// TwinCAT 3 PLC project PLC
// ProgramVersion: 3.1.4026.28
// libraries:
//   Tc2_MC2, * (Beckhoff Automation GmbH)
//   Tc2_Standard, * (Beckhoff Automation GmbH)
//   Tc2_System, * (Beckhoff Automation GmbH)
// project tree:
//   Adapters/Nc/ Axes.TcGVL, DriveAxis_Nc.TcPOU
//   Adapters/Simulation/ Accelerometer_Simulated.TcPOU, DigitalOut_SimulatedLidarPower.TcPOU, Gyro_Simulated.TcPOU, Lidar_Simulated.TcPOU, SimulatorLink.TcPOU
//   App/ MAIN.TcPOU, RobotComposition.TcPOU
//   Contracts/ HmiCommand.TcDUT, HmiCommandCode.TcDUT, HmiStatus.TcDUT, MapInfo.TcDUT, MissionState.TcDUT, RobotHmi.TcGVL, SimulatorCommand.TcDUT, SimulatorFeedback.TcDUT, SimulatorIo.TcGVL
//   Core/ BodyMotion.TcDUT, Constants.TcGVL, HardwareError.TcDUT, LaserScan.TcDUT, Parameters.TcGVL, PlatformKind.TcDUT, Pose2D.TcDUT, Twist.TcDUT, Vector3.TcDUT, WheelSpeeds.TcDUT
//   Hal/ I_Accelerometer.TcIO, I_DigitalOut.TcIO, I_DriveAxis.TcIO, I_Gyro.TcIO, I_Lidar.TcIO, Lidar_Watchdog.TcPOU
//   Localization/ I_PoseSource.TcIO, GyroOdometry.TcPOU, WheelOdometry.TcPOU
//   Mapping/ GridCell.TcDUT, OccupancyGrid.TcPOU
//   Mission/ SweepMission.TcPOU
//   Platform/ DiffDrive.TcPOU, DiffDriveKinematics.TcPOU, I_DifferentialDrive.TcIO
//   / PlcTask.TcTTO
// real-time tasks:
//   TASK PlcTask: cycle T#10ms, priority 20, ADS port 350
// motion (NC):
//   TASK NC-Task 1 SAF: cycle T#2ms, priority 4, ADS port 501
//   TASK NC-Task 1 SVB: cycle T#10ms, priority 8, ADS port 511
//   AXIS LeftWheel (id 1)
//     General: UnitName=m
//     Dynamic: AccelerationMaximum=2, DecelerationMaximum=2, Acceleration=1, Deceleration=1, Jerk=10
//     Velo: Maximum=0.6
//     OtherSettings: AllowMotionCmdToSlave=true
//     encoder EncType=1
//     drive DrvType=5
//       Analog: VeloReferenz=0.6, TorqueSetpointScale=10, ScaleFactorActTorque=0.1
//       TimeComp: TaskDelayCycles=1
//     controller CtrType=1
//       CtrPara: PriorControlFactor=1
//         Observer: BandWidth=20
//   AXIS RightWheel (id 2)
//     General: UnitName=m
//     Dynamic: AccelerationMaximum=2, DecelerationMaximum=2, Acceleration=1, Deceleration=1, Jerk=10
//     Velo: Maximum=0.6
//     OtherSettings: AllowMotionCmdToSlave=true
//     encoder EncType=1
//     drive DrvType=5
//       Analog: VeloReferenz=0.6, TorqueSetpointScale=10, ScaleFactorActTorque=0.1
//       TimeComp: TaskDelayCycles=1
//     controller CtrType=1
//       CtrPara: PriorControlFactor=1
//         Observer: BandWidth=20
// variable links:
//   PLC/PLC Instance <-> NC-Task 1 SAF/Axes/LeftWheel
//     PlcTask Inputs/Axes.leftWheel.NcToPlc <-> Outputs/ToPlc
//     PlcTask Outputs/Axes.leftWheel.PlcToNc <-> Inputs/FromPlc
//   PLC/PLC Instance <-> NC-Task 1 SAF/Axes/RightWheel
//     PlcTask Inputs/Axes.rightWheel.NcToPlc <-> Outputs/ToPlc
//     PlcTask Outputs/Axes.rightWheel.PlcToNc <-> Inputs/FromPlc

CONFIGURATION PLC
    RESOURCE PLC ON TwinCAT3
        TASK PlcTask(INTERVAL := T#10ms, PRIORITY := 20);
        PROGRAM MAIN WITH PlcTask : MAIN;
    END_RESOURCE
END_CONFIGURATION

// ---- Contracts/HmiCommand.TcDUT
TYPE HmiCommand :
STRUCT
	sequence : UDINT;
	code : HmiCommandCode;
	manualTwist : Twist;
	pose : Pose2D;
END_STRUCT
END_TYPE

// ---- Contracts/HmiCommandCode.TcDUT
{attribute 'qualified_only'}
{attribute 'strict'}
TYPE HmiCommandCode :
(
	NONE := 0,
	MANUAL_DRIVE,
	START_MAPPING,
	START_SWEEPING,
	PAUSE,
	RESUME,
	STOP,
	GO_TO_DOCK,
	EMERGENCY_STOP,
	RESET,
	SET_POSE
) INT;
END_TYPE

// ---- Contracts/HmiStatus.TcDUT
TYPE HmiStatus :
STRUCT
	acknowledgedSequence : UDINT;
	missionState : MissionState;
	lastRejection : STRING(80);
	estimatedPose : Pose2D;
	isSimulatorConnected : BOOL;
	isLidarOk : BOOL;
	hasMap : BOOL;
END_STRUCT
END_TYPE

// ---- Contracts/MapInfo.TcDUT
// Det GUI-en trenger for å tegne RobotHmi.mapCells.
TYPE MapInfo :
STRUCT
	// Øker hver gang kartet er endret, så serveren bare henter cellene på nytt når det trengs.
	revision : UDINT;
	cellSizeInM : LREAL;
	// Hjørnet til celle [0, 0] i verden.
	originXInM : LREAL;
	originYInM : LREAL;
	widthInCells : UINT;
	heightInCells : UINT;
	// Hvor mye log-odds én enhet i en celle er. 0.1 betyr at 35 i cella er log-odds 3.5.
	logOddsPerUnit : LREAL;
END_STRUCT
END_TYPE

// ---- Contracts/MissionState.TcDUT
{attribute 'qualified_only'}
{attribute 'strict'}
TYPE MissionState :
(
	IDLE := 0,
	MANUAL,
	MAPPING,
	SWEEPING,
	PAUSED,
	RETURNING_TO_DOCK,
	DOCKED,
	EMERGENCY_STOPPED
) INT;
END_TYPE

// ---- Contracts/SimulatorCommand.TcDUT
TYPE SimulatorCommand :
STRUCT
	version : UDINT;
	cycle : UDINT;
	plcTimeInNs : ULINT;
	// The wheels' actual speed and position, from the NC axes. The simulated wheels run at
	// the speed and are nudged towards the position, so they never drift away from NC.
	leftWheelVelocityInMPerS : LREAL;
	rightWheelVelocityInMPerS : LREAL;
	leftWheelPositionInM : LREAL;
	rightWheelPositionInM : LREAL;
	isLeftDriveEnabled : BOOL;
	isRightDriveEnabled : BOOL;
	isLidarPowered : BOOL;
	estimatedPose : Pose2D;
END_STRUCT
END_TYPE

// ---- Contracts/SimulatorFeedback.TcDUT
TYPE SimulatorFeedback :
STRUCT
	version : UDINT;
	sequence : UDINT;
	timeInNs : ULINT;
	leftWheelAngleInRad : LREAL;
	rightWheelAngleInRad : LREAL;
	leftWheelVelocityInRadPerS : LREAL;
	rightWheelVelocityInRadPerS : LREAL;
	angularRateInRadPerS : Vector3;
	accelerationInMPerS2 : Vector3;
	truePose : Pose2D;
	collided : BOOL;
END_STRUCT
END_TYPE

// ---- Core/BodyMotion.TcDUT
TYPE BodyMotion :
STRUCT
	distanceInM : LREAL;
	headingChangeInRad : LREAL;
END_STRUCT
END_TYPE

// ---- Core/HardwareError.TcDUT
TYPE HardwareError :
STRUCT
	isActive : BOOL;
	id : UDINT;
	text : STRING(80);
END_STRUCT
END_TYPE

// ---- Core/LaserScan.TcDUT
TYPE LaserScan :
STRUCT
	sequence : UDINT;
	startTimestampInNs : ULINT;
	scanDurationInS : REAL;
	angleMinInRad : REAL;
	angleIncrementInRad : REAL;
	count : UINT;
	rangesInM : ARRAY[0..Constants.MAX_SCAN_POINTS - 1] OF REAL;
END_STRUCT
END_TYPE

// ---- Core/PlatformKind.TcDUT
{attribute 'qualified_only'}
{attribute 'strict'}
TYPE PlatformKind :
(
	SIMULATION := 0,
	HARDWARE
);
END_TYPE

// ---- Core/Pose2D.TcDUT
TYPE Pose2D :
STRUCT
	x : LREAL;
	y : LREAL;
	thetaInRad : LREAL;
END_STRUCT
END_TYPE

// ---- Core/Twist.TcDUT
TYPE Twist :
STRUCT
	forwardSpeedInMPerS : LREAL;
	yawRateInRadPerS : LREAL;
END_STRUCT
END_TYPE

// ---- Core/Vector3.TcDUT
TYPE Vector3 :
STRUCT
	x : LREAL;
	y : LREAL;
	z : LREAL;
END_STRUCT
END_TYPE

// ---- Core/WheelSpeeds.TcDUT
TYPE WheelSpeeds :
STRUCT
	leftInMPerS : LREAL;
	rightInMPerS : LREAL;
END_STRUCT
END_TYPE

// ---- Mapping/GridCell.TcDUT
// Én rute i kartet. x teller østover og y nordover fra kartets origo, som i verden.
TYPE GridCell :
STRUCT
	x : DINT;
	y : DINT;
END_STRUCT
END_TYPE

// ---- Adapters/Nc/Axes.TcGVL
{attribute 'qualified_only'}
VAR_GLOBAL
	// Link each one to its NC axis in XAE: the axis, Settings, Link To PLC.
	leftWheel : AXIS_REF;
	rightWheel : AXIS_REF;
END_VAR

// ---- Contracts/RobotHmi.TcGVL
{attribute 'qualified_only'}
VAR_GLOBAL
	command : HmiCommand;
	status : HmiStatus;
	// Kartet PLC-en bygger, for GUI-en. Indeksen er [x, y]; y endrer seg raskest i minnet.
	mapInfo : MapInfo;
	mapCells : ARRAY[0..Constants.MAP_WIDTH_IN_CELLS - 1, 0..Constants.MAP_HEIGHT_IN_CELLS - 1] OF SINT;
END_VAR

// ---- Contracts/SimulatorIo.TcGVL
{attribute 'qualified_only'}
VAR_GLOBAL
	command : SimulatorCommand;
	feedback : SimulatorFeedback;
	scan : LaserScan;
END_VAR

// ---- Core/Constants.TcGVL
{attribute 'qualified_only'}
VAR_GLOBAL CONSTANT
	MAX_SCAN_POINTS : UINT := 1024;
	// Kartet er 256 x 256 ruter. Med 5 cm ruter blir det 12,8 x 12,8 m.
	MAP_WIDTH_IN_CELLS : UINT := 256;
	MAP_HEIGHT_IN_CELLS : UINT := 256;
	// Én enhet i en kartcelle er så mye log-odds.
	MAP_LOG_ODDS_PER_UNIT : LREAL := 0.1;
	SIMULATOR_PROTOCOL_VERSION : UDINT := 4;
	SIMULATOR_TIMEOUT_IN_CYCLES : UDINT := 20;
	LIDAR_TIMEOUT_IN_MS : TIME := T#400MS;
	SIMULATOR_NOT_CONNECTED_ERROR_ID : UDINT := 1001;
	LIDAR_TIMEOUT_ERROR_ID : UDINT := 2001;
	AXIS_NOT_LINKED_ERROR_ID : UDINT := 3001;
END_VAR

// ---- Core/Parameters.TcGVL
{attribute 'qualified_only'}
VAR_GLOBAL PERSISTENT
	platform : PlatformKind := PlatformKind.SIMULATION;
	// Hjulradien ligger i NC-skaleringen av aksene, som går i meter langs hjulbanen.
	trackWidthInM : LREAL := 0.40;
	maxWheelSpeedInMPerS : LREAL := 0.6;
	// Hvor fort hjulene får endre fart. Uten disse bruker NC sine standardverdier, og hjulene
	// stopper fra full fart på et par hundredeler, mye brattere enn en ekte robot tåler uten å skli.
	wheelAccelerationInMPerS2 : LREAL := 1.0;
	wheelJerkInMPerS3 : LREAL := 10.0;
	useGyroForHeading : BOOL := FALSE;
	gyroScale : LREAL := 1.0;

	// Hvor lidaren sitter på roboten, sett fra midt mellom hjulene (x fram, y mot venstre),
	// og hvor mye den er dreid. I simulatoren står den midt mellom hjulene og peker rett fram.
	lidarMountXInM : LREAL := 0.0;
	lidarMountYInM : LREAL := 0.0;
	lidarMountThetaInRad : LREAL := 0.0;

	// Kartet. Origo er hjørnet til celle [0, 0]; med -3.4 dekker kartet en garasje på 6 x 6 m med god margin.
	mapCellSizeInM : LREAL := 0.05;
	mapOriginXInM : LREAL := -3.4;
	mapOriginYInM : LREAL := -3.4;
	// Log-odds i tideler (Constants.MAP_LOG_ODDS_PER_UNIT): treff +0.9, fri -0.4, aldri mer enn ±3.5.
	mapHitLogOdds : SINT := 9;
	mapFreeLogOdds : SINT := -4;
	mapMaxLogOdds : SINT := 35;
END_VAR

// ---- Hal/I_Accelerometer.TcIO
INTERFACE I_Accelerometer

PROPERTY AccelerationInMPerS2 : Vector3
GET
END_GET
END_PROPERTY

PROPERTY TimestampInNs : ULINT
GET
END_GET
END_PROPERTY

PROPERTY IsValid : BOOL
GET
END_GET
END_PROPERTY

END_INTERFACE

// ---- Hal/I_DigitalOut.TcIO
INTERFACE I_DigitalOut

METHOD SwitchOn
END_METHOD

METHOD SwitchOff
END_METHOD

PROPERTY IsOn : BOOL
GET
END_GET
END_PROPERTY

END_INTERFACE

// ---- Hal/I_DriveAxis.TcIO
INTERFACE I_DriveAxis

METHOD Execute
END_METHOD

METHOD Enable
END_METHOD

METHOD Disable
END_METHOD

METHOD SetVelocity
VAR_INPUT
	velocityInMPerS : LREAL;
END_VAR
END_METHOD

METHOD TryReset : BOOL
END_METHOD

PROPERTY PositionInM : LREAL
GET
END_GET
END_PROPERTY

PROPERTY VelocityInMPerS : LREAL
GET
END_GET
END_PROPERTY

PROPERTY IsReady : BOOL
GET
END_GET
END_PROPERTY

PROPERTY IsStandingStill : BOOL
GET
END_GET
END_PROPERTY

PROPERTY Error : HardwareError
GET
END_GET
END_PROPERTY

END_INTERFACE

// ---- Hal/I_Gyro.TcIO
INTERFACE I_Gyro

METHOD StartBiasCalibration
END_METHOD

PROPERTY YawRateInRadPerS : LREAL
GET
END_GET
END_PROPERTY

PROPERTY AngularRateInRadPerS : Vector3
GET
END_GET
END_PROPERTY

PROPERTY TimestampInNs : ULINT
GET
END_GET
END_PROPERTY

PROPERTY IsValid : BOOL
GET
END_GET
END_PROPERTY

END_INTERFACE

// ---- Hal/I_Lidar.TcIO
INTERFACE I_Lidar

METHOD Start
END_METHOD

METHOD Stop
END_METHOD

METHOD TryGetScan : BOOL
VAR_INPUT
	scan : REFERENCE TO LaserScan;
END_VAR
END_METHOD

PROPERTY IsRunning : BOOL
GET
END_GET
END_PROPERTY

PROPERTY Error : HardwareError
GET
END_GET
END_PROPERTY

END_INTERFACE

// ---- Localization/I_PoseSource.TcIO
INTERFACE I_PoseSource

METHOD Reset
VAR_INPUT
	pose : Pose2D;
END_VAR
END_METHOD

PROPERTY Pose : Pose2D
GET
END_GET
END_PROPERTY

END_INTERFACE

// ---- Platform/I_DifferentialDrive.TcIO
INTERFACE I_DifferentialDrive

METHOD Execute
END_METHOD

METHOD Enable
END_METHOD

METHOD Disable
END_METHOD

METHOD SetTwist
VAR_INPUT
	desiredTwist : Twist;
END_VAR
END_METHOD

PROPERTY LeftWheelPositionInM : LREAL
GET
END_GET
END_PROPERTY

PROPERTY RightWheelPositionInM : LREAL
GET
END_GET
END_PROPERTY

PROPERTY IsReady : BOOL
GET
END_GET
END_PROPERTY

PROPERTY IsStandingStill : BOOL
GET
END_GET
END_PROPERTY

END_INTERFACE

// ---- App/MAIN.TcPOU
PROGRAM MAIN
VAR
	robot : RobotComposition;
END_VAR

robot.Execute();

END_PROGRAM

// ---- App/RobotComposition.TcPOU
{attribute 'linkalways'}
{attribute 'no_explicit_call' := 'Use the methods of this class'}
{attribute 'enable_dynamic_creation'}
FUNCTION_BLOCK RobotComposition
VAR
	simulator : SimulatorLink;
	leftAxis : DriveAxis_Nc(ncAxis := Axes.leftWheel);
	rightAxis : DriveAxis_Nc(ncAxis := Axes.rightWheel);
	simulatedGyro : Gyro_Simulated(simulator := simulator);
	simulatedAccelerometer : Accelerometer_Simulated(simulator := simulator);
	simulatedLidar : Lidar_Simulated(simulator := simulator);
	simulatedLidarPower : DigitalOut_SimulatedLidarPower;

	gyro : I_Gyro;
	accelerometer : I_Accelerometer;
	lidarPower : I_DigitalOut;
	lidar : Lidar_Watchdog;
	drive : DiffDrive;
	odometry : WheelOdometry;
	gyroOdometry : GyroOdometry;
	grid : OccupancyGrid;
	mission : SweepMission;

	scan : LaserScan;
	requestedPose : Pose2D;
	isInitialized : BOOL;
END_VAR

METHOD Execute
IF NOT isInitialized THEN
	Initialize();
END_IF

IF Parameters.platform = PlatformKind.SIMULATION THEN
	simulator.Execute();
END_IF

lidar.Execute();
IF lidar.TryGetScan(scan) AND mission.State = MissionState.MAPPING THEN
	// Kommer i M4: scan matching, som retter posisjonen mot kartet før scannet legges inn.
	grid.Integrate(scan := scan, pose := EstimatedPose());
	grid.Publish(RobotHmi.mapInfo, RobotHmi.mapCells);
END_IF

odometry.Execute();
gyroOdometry.Execute();
mission.Execute();
IF mission.TryTakePoseRequest(requestedPose) THEN
	odometry.Reset(requestedPose);
	gyroOdometry.Reset(requestedPose);
END_IF
IF mission.TryTakeMapClearRequest() THEN
	grid.Clear();
	grid.Publish(RobotHmi.mapInfo, RobotHmi.mapCells);
END_IF

IF mission.ShouldDrive THEN
	drive.Enable();
	drive.SetTwist(mission.DesiredTwist);
ELSE
	drive.Disable();
END_IF
drive.Execute();

IF Parameters.platform = PlatformKind.SIMULATION THEN
	SendWheelsToSimulator();
END_IF

PublishStatus();
END_METHOD

METHOD PRIVATE Initialize
VAR
	start : Pose2D;
END_VAR
CASE Parameters.platform OF
	PlatformKind.SIMULATION:
		gyro := simulatedGyro;
		accelerometer := simulatedAccelerometer;
		lidar.Wrap(simulatedLidar);
		lidarPower := simulatedLidarPower;
	PlatformKind.HARDWARE:
		// Kommer i M7: Gyro_EP3751 og valgt LIDAR-adapter. Hjulene bruker de samme NC-aksene.
		RETURN;
END_CASE

drive.Connect(leftAxis, rightAxis);

lidarPower.SwitchOn();
lidar.Start();
odometry.Connect(drive);
odometry.Reset(start);
gyroOdometry.Connect(drive, gyro);
gyroOdometry.Reset(start);
grid.Clear();
grid.Publish(RobotHmi.mapInfo, RobotHmi.mapCells);
isInitialized := TRUE;
END_METHOD

METHOD PRIVATE SendWheelsToSimulator
// I simuleringen er NC-aksene motor og enkoder. Simulatoren får vite hvor langt hjulene faktisk har gått,
// lar de simulerte hjulene følge det nøyaktig, og flytter roboten etter det, med sluring og kollisjoner.
SimulatorIo.command.leftWheelVelocityInMPerS := leftAxis.VelocityInMPerS;
SimulatorIo.command.rightWheelVelocityInMPerS := rightAxis.VelocityInMPerS;
SimulatorIo.command.leftWheelPositionInM := leftAxis.PositionInM;
SimulatorIo.command.rightWheelPositionInM := rightAxis.PositionInM;
SimulatorIo.command.isLeftDriveEnabled := leftAxis.IsReady;
SimulatorIo.command.isRightDriveEnabled := rightAxis.IsReady;
END_METHOD

METHOD PRIVATE PublishStatus
VAR
	lidarError : HardwareError;
	estimate : Pose2D;
END_VAR
estimate := EstimatedPose();
lidarError := lidar.Error;
RobotHmi.status.estimatedPose := estimate;
RobotHmi.status.isSimulatorConnected := simulator.IsConnected;
RobotHmi.status.isLidarOk := NOT lidarError.isActive;
SimulatorIo.command.estimatedPose := estimate;
END_METHOD

// Den posisjonen roboten tror den har, fra estimatet Parameters.useGyroForHeading velger.
METHOD PRIVATE EstimatedPose : Pose2D
IF Parameters.useGyroForHeading THEN
	EstimatedPose := gyroOdometry.Pose;
ELSE
	EstimatedPose := odometry.Pose;
END_IF
END_METHOD

END_FUNCTION_BLOCK

// ---- Adapters/Simulation/SimulatorLink.TcPOU
{attribute 'linkalways'}
{attribute 'no_explicit_call' := 'Use the methods of this class'}
{attribute 'enable_dynamic_creation'}
FUNCTION_BLOCK SimulatorLink
VAR
	cycle : UDINT;
	lastSequence : UDINT;
	silentCycles : UDINT;
	_isConnected : BOOL;
END_VAR

METHOD Execute
cycle := cycle + 1;
SimulatorIo.command.version := Constants.SIMULATOR_PROTOCOL_VERSION;
SimulatorIo.command.cycle := cycle;
SimulatorIo.command.plcTimeInNs := F_GetSystemTime() * 100;

IF SimulatorIo.feedback.sequence <> lastSequence THEN
	lastSequence := SimulatorIo.feedback.sequence;
	silentCycles := 0;
ELSIF silentCycles < Constants.SIMULATOR_TIMEOUT_IN_CYCLES THEN
	silentCycles := silentCycles + 1;
END_IF

_isConnected := SimulatorIo.feedback.version = Constants.SIMULATOR_PROTOCOL_VERSION
	AND silentCycles < Constants.SIMULATOR_TIMEOUT_IN_CYCLES;
END_METHOD

PROPERTY IsConnected : BOOL
GET
IsConnected := _isConnected;
END_GET
END_PROPERTY

END_FUNCTION_BLOCK

// ---- Adapters/Nc/DriveAxis_Nc.TcPOU
{attribute 'linkalways'}
{attribute 'no_explicit_call' := 'Use the methods of this class'}
{attribute 'enable_dynamic_creation'}
FUNCTION_BLOCK DriveAxis_Nc IMPLEMENTS I_DriveAxis
VAR
	axis : REFERENCE TO AXIS_REF;
	power : MC_Power;
	moveVelocity : MC_MoveVelocity;
	halt : MC_Halt;
	reset : MC_Reset;
	isEnabled : BOOL;
	targetInMPerS : LREAL;
	commandedInMPerS : LREAL;
	isHalting : BOOL;
	notLinkedError : HardwareError := (isActive := TRUE, id := Constants.AXIS_NOT_LINKED_ERROR_ID, text := 'Aksen er ikke koblet til PLC-en');
END_VAR
VAR CONSTANT
	// NC refuses set velocities below 0.001 (axis unit/s), so anything slower is a stop.
	MIN_VELOCITY_IN_M_PER_S : LREAL := 0.001;
	VELOCITY_DEADBAND_IN_M_PER_S : LREAL := 0.0005;
END_VAR

METHOD FB_init : BOOL
VAR_INPUT
	bInitRetains : BOOL;
	bInCopyCode : BOOL;
	ncAxis : REFERENCE TO AXIS_REF;
END_VAR
axis REF= ncAxis;
END_METHOD

METHOD Execute
IF NOT __ISVALIDREF(axis) THEN
	RETURN;
END_IF
axis.ReadStatus();
power(Axis := axis, Enable := isEnabled, Enable_Positive := isEnabled, Enable_Negative := isEnabled, Override := 100);
reset(Axis := axis, Execute := FALSE);

IF NOT isEnabled OR NOT power.Status THEN
	commandedInMPerS := 0;
	isHalting := FALSE;
	moveVelocity(Axis := axis, Execute := FALSE);
	halt(Axis := axis, Execute := FALSE);
	RETURN;
END_IF

IF ABS(targetInMPerS) < MIN_VELOCITY_IN_M_PER_S THEN
	IF NOT isHalting THEN
		isHalting := TRUE;
		commandedInMPerS := 0;
		moveVelocity(Axis := axis, Execute := FALSE);
		halt(Axis := axis, Execute := FALSE);
	END_IF
	halt(
		Axis := axis,
		Execute := TRUE,
		Deceleration := Parameters.wheelAccelerationInMPerS2,
		Jerk := Parameters.wheelJerkInMPerS3);
ELSIF isHalting OR ABS(targetInMPerS - commandedInMPerS) > VELOCITY_DEADBAND_IN_M_PER_S THEN
	// MC_MoveVelocity starts on a rising edge, so a new speed needs Execute low, then high.
	isHalting := FALSE;
	commandedInMPerS := targetInMPerS;
	halt(Axis := axis, Execute := FALSE);
	moveVelocity(Axis := axis, Execute := FALSE);
	moveVelocity(
		Axis := axis,
		Execute := TRUE,
		Velocity := ABS(targetInMPerS),
		Acceleration := Parameters.wheelAccelerationInMPerS2,
		Deceleration := Parameters.wheelAccelerationInMPerS2,
		Jerk := Parameters.wheelJerkInMPerS3,
		Direction := SEL(targetInMPerS > 0, MC_Negative_Direction, MC_Positive_Direction));
ELSE
	moveVelocity(Axis := axis, Execute := TRUE);
END_IF
END_METHOD

METHOD Enable
isEnabled := TRUE;
END_METHOD

METHOD Disable
isEnabled := FALSE;
targetInMPerS := 0;
END_METHOD

METHOD SetVelocity
VAR_INPUT
	velocityInMPerS : LREAL;
END_VAR
targetInMPerS := LIMIT(-Parameters.maxWheelSpeedInMPerS, velocityInMPerS, Parameters.maxWheelSpeedInMPerS);
END_METHOD

METHOD TryReset : BOOL
IF NOT __ISVALIDREF(axis) THEN
	RETURN;
END_IF
reset(Axis := axis, Execute := TRUE);
TryReset := NOT axis.Status.Error;
END_METHOD

PROPERTY PositionInM : LREAL
GET
IF __ISVALIDREF(axis) THEN
	PositionInM := axis.NcToPlc.ActPos;
END_IF
END_GET
END_PROPERTY

PROPERTY VelocityInMPerS : LREAL
GET
IF __ISVALIDREF(axis) THEN
	VelocityInMPerS := axis.NcToPlc.ActVelo;
END_IF
END_GET
END_PROPERTY

PROPERTY IsReady : BOOL
GET
IsReady := __ISVALIDREF(axis) AND_THEN power.Status AND NOT axis.Status.Error;
END_GET
END_PROPERTY

PROPERTY IsStandingStill : BOOL
GET
IsStandingStill := __ISVALIDREF(axis) AND_THEN axis.Status.NotMoving;
END_GET
END_PROPERTY

PROPERTY Error : HardwareError
GET
VAR
	axisError : HardwareError;
END_VAR
IF NOT __ISVALIDREF(axis) THEN
	Error := notLinkedError;
ELSIF axis.Status.Error THEN
	axisError.isActive := TRUE;
	axisError.id := axis.Status.ErrorID;
	axisError.text := 'NC-aksen melder feil, se feilkoden';
	Error := axisError;
END_IF
END_GET
END_PROPERTY

END_FUNCTION_BLOCK

// ---- Adapters/Simulation/Gyro_Simulated.TcPOU
{attribute 'linkalways'}
{attribute 'no_explicit_call' := 'Use the methods of this class'}
{attribute 'enable_dynamic_creation'}
FUNCTION_BLOCK Gyro_Simulated IMPLEMENTS I_Gyro
VAR
	link : REFERENCE TO SimulatorLink;
END_VAR

METHOD FB_init : BOOL
VAR_INPUT
	bInitRetains : BOOL;
	bInCopyCode : BOOL;
	simulator : REFERENCE TO SimulatorLink;
END_VAR
link REF= simulator;
END_METHOD

METHOD StartBiasCalibration
// The simulated gyro has no calibration of its own. Bias is estimated in GyroOdometry.
END_METHOD

PROPERTY YawRateInRadPerS : LREAL
GET
YawRateInRadPerS := SimulatorIo.feedback.angularRateInRadPerS.z;
END_GET
END_PROPERTY

PROPERTY AngularRateInRadPerS : Vector3
GET
AngularRateInRadPerS := SimulatorIo.feedback.angularRateInRadPerS;
END_GET
END_PROPERTY

PROPERTY TimestampInNs : ULINT
GET
TimestampInNs := SimulatorIo.feedback.timeInNs;
END_GET
END_PROPERTY

PROPERTY IsValid : BOOL
GET
IsValid := __ISVALIDREF(link) AND_THEN link.IsConnected;
END_GET
END_PROPERTY

END_FUNCTION_BLOCK

// ---- Adapters/Simulation/Accelerometer_Simulated.TcPOU
{attribute 'linkalways'}
{attribute 'no_explicit_call' := 'Use the methods of this class'}
{attribute 'enable_dynamic_creation'}
FUNCTION_BLOCK Accelerometer_Simulated IMPLEMENTS I_Accelerometer
VAR
	link : REFERENCE TO SimulatorLink;
END_VAR

METHOD FB_init : BOOL
VAR_INPUT
	bInitRetains : BOOL;
	bInCopyCode : BOOL;
	simulator : REFERENCE TO SimulatorLink;
END_VAR
link REF= simulator;
END_METHOD

PROPERTY AccelerationInMPerS2 : Vector3
GET
AccelerationInMPerS2 := SimulatorIo.feedback.accelerationInMPerS2;
END_GET
END_PROPERTY

PROPERTY TimestampInNs : ULINT
GET
TimestampInNs := SimulatorIo.feedback.timeInNs;
END_GET
END_PROPERTY

PROPERTY IsValid : BOOL
GET
IsValid := __ISVALIDREF(link) AND_THEN link.IsConnected;
END_GET
END_PROPERTY

END_FUNCTION_BLOCK

// ---- Adapters/Simulation/Lidar_Simulated.TcPOU
{attribute 'linkalways'}
{attribute 'no_explicit_call' := 'Use the methods of this class'}
{attribute 'enable_dynamic_creation'}
FUNCTION_BLOCK Lidar_Simulated IMPLEMENTS I_Lidar
VAR
	notConnectedError : HardwareError := (isActive := TRUE, id := Constants.SIMULATOR_NOT_CONNECTED_ERROR_ID, text := 'Simulatoren er ikke tilkoblet');
	link : REFERENCE TO SimulatorLink;
	_isRunning : BOOL;
	lastSequence : UDINT;
END_VAR

METHOD FB_init : BOOL
VAR_INPUT
	bInitRetains : BOOL;
	bInCopyCode : BOOL;
	simulator : REFERENCE TO SimulatorLink;
END_VAR
link REF= simulator;
END_METHOD

METHOD Start
_isRunning := TRUE;
lastSequence := SimulatorIo.scan.sequence;
END_METHOD

METHOD Stop
_isRunning := FALSE;
END_METHOD

METHOD TryGetScan : BOOL
VAR_INPUT
	scan : REFERENCE TO LaserScan;
END_VAR
IF NOT _isRunning OR_ELSE SimulatorIo.scan.sequence = lastSequence THEN
	RETURN;
END_IF
lastSequence := SimulatorIo.scan.sequence;
scan := SimulatorIo.scan;
TryGetScan := TRUE;
END_METHOD

PROPERTY IsRunning : BOOL
GET
IsRunning := _isRunning;
END_GET
END_PROPERTY

PROPERTY Error : HardwareError
GET
IF NOT __ISVALIDREF(link) OR_ELSE NOT link.IsConnected THEN
	Error := notConnectedError;
END_IF
END_GET
END_PROPERTY

END_FUNCTION_BLOCK

// ---- Adapters/Simulation/DigitalOut_SimulatedLidarPower.TcPOU
{attribute 'linkalways'}
{attribute 'no_explicit_call' := 'Use the methods of this class'}
{attribute 'enable_dynamic_creation'}
FUNCTION_BLOCK DigitalOut_SimulatedLidarPower IMPLEMENTS I_DigitalOut

METHOD SwitchOn
SimulatorIo.command.isLidarPowered := TRUE;
END_METHOD

METHOD SwitchOff
SimulatorIo.command.isLidarPowered := FALSE;
END_METHOD

PROPERTY IsOn : BOOL
GET
IsOn := SimulatorIo.command.isLidarPowered;
END_GET
END_PROPERTY

END_FUNCTION_BLOCK

// ---- Hal/Lidar_Watchdog.TcPOU
{attribute 'linkalways'}
{attribute 'no_explicit_call' := 'Use the methods of this class'}
{attribute 'enable_dynamic_creation'}
FUNCTION_BLOCK Lidar_Watchdog IMPLEMENTS I_Lidar
VAR
	timeoutError : HardwareError := (isActive := TRUE, id := Constants.LIDAR_TIMEOUT_ERROR_ID, text := 'Ingen LIDAR-skann innenfor fristen');
	inner : I_Lidar;
	timeoutTimer : TON;
	isTimedOut : BOOL;
END_VAR

METHOD Wrap
VAR_INPUT
	lidar : I_Lidar;
END_VAR
inner := lidar;
END_METHOD

METHOD Execute
IF inner = 0 THEN
	RETURN;
END_IF
timeoutTimer(IN := inner.IsRunning, PT := Constants.LIDAR_TIMEOUT_IN_MS);
IF timeoutTimer.Q THEN
	isTimedOut := TRUE;
END_IF
END_METHOD

METHOD Start
IF inner <> 0 THEN
	inner.Start();
END_IF
timeoutTimer(IN := FALSE);
isTimedOut := FALSE;
END_METHOD

METHOD Stop
IF inner <> 0 THEN
	inner.Stop();
END_IF
timeoutTimer(IN := FALSE);
isTimedOut := FALSE;
END_METHOD

METHOD TryGetScan : BOOL
VAR_INPUT
	scan : REFERENCE TO LaserScan;
END_VAR
IF inner = 0 OR_ELSE NOT inner.TryGetScan(scan) THEN
	RETURN;
END_IF
timeoutTimer(IN := FALSE);
isTimedOut := FALSE;
TryGetScan := TRUE;
END_METHOD

PROPERTY IsRunning : BOOL
GET
IsRunning := inner <> 0 AND_THEN inner.IsRunning;
END_GET
END_PROPERTY

PROPERTY Error : HardwareError
GET
IF isTimedOut THEN
	Error := timeoutError;
ELSIF inner <> 0 THEN
	Error := inner.Error;
END_IF
END_GET
END_PROPERTY

END_FUNCTION_BLOCK

// ---- Platform/DiffDrive.TcPOU
{attribute 'linkalways'}
{attribute 'no_explicit_call' := 'Use the methods of this class'}
{attribute 'enable_dynamic_creation'}
FUNCTION_BLOCK DiffDrive IMPLEMENTS I_DifferentialDrive
VAR
	leftAxis : I_DriveAxis;
	rightAxis : I_DriveAxis;
	kinematics : DiffDriveKinematics;
END_VAR

METHOD Connect
VAR_INPUT
	left : I_DriveAxis;
	right : I_DriveAxis;
END_VAR
leftAxis := left;
rightAxis := right;
END_METHOD

METHOD Execute
IF leftAxis = 0 OR rightAxis = 0 THEN
	RETURN;
END_IF
leftAxis.Execute();
rightAxis.Execute();
END_METHOD

METHOD Enable
IF leftAxis = 0 OR rightAxis = 0 THEN
	RETURN;
END_IF
leftAxis.Enable();
rightAxis.Enable();
END_METHOD

METHOD Disable
IF leftAxis = 0 OR rightAxis = 0 THEN
	RETURN;
END_IF
leftAxis.Disable();
rightAxis.Disable();
END_METHOD

METHOD SetTwist
VAR_INPUT
	desiredTwist : Twist;
END_VAR
VAR
	speeds : WheelSpeeds;
END_VAR
IF leftAxis = 0 OR rightAxis = 0 THEN
	RETURN;
END_IF
speeds := kinematics.ToWheelSpeeds(desiredTwist);
leftAxis.SetVelocity(speeds.leftInMPerS);
rightAxis.SetVelocity(speeds.rightInMPerS);
END_METHOD

PROPERTY LeftWheelPositionInM : LREAL
GET
IF leftAxis <> 0 THEN
	LeftWheelPositionInM := leftAxis.PositionInM;
END_IF
END_GET
END_PROPERTY

PROPERTY RightWheelPositionInM : LREAL
GET
IF rightAxis <> 0 THEN
	RightWheelPositionInM := rightAxis.PositionInM;
END_IF
END_GET
END_PROPERTY

PROPERTY IsReady : BOOL
GET
IsReady := leftAxis <> 0 AND_THEN rightAxis <> 0 AND_THEN leftAxis.IsReady AND_THEN rightAxis.IsReady;
END_GET
END_PROPERTY

PROPERTY IsStandingStill : BOOL
GET
IsStandingStill := leftAxis <> 0 AND_THEN rightAxis <> 0 AND_THEN leftAxis.IsStandingStill AND_THEN rightAxis.IsStandingStill;
END_GET
END_PROPERTY

END_FUNCTION_BLOCK

// ---- Platform/DiffDriveKinematics.TcPOU
{attribute 'linkalways'}
{attribute 'no_explicit_call' := 'Use the methods of this class'}
{attribute 'enable_dynamic_creation'}
FUNCTION_BLOCK DiffDriveKinematics

METHOD ToBodyMotion : BodyMotion
VAR_INPUT
	leftDeltaInM : LREAL;
	rightDeltaInM : LREAL;
END_VAR
VAR
	motion : BodyMotion;
END_VAR
motion.distanceInM := (leftDeltaInM + rightDeltaInM) / 2.0;
motion.headingChangeInRad := (rightDeltaInM - leftDeltaInM) / Parameters.trackWidthInM;

ToBodyMotion := motion;
END_METHOD

METHOD ToWheelSpeeds : WheelSpeeds
VAR_INPUT
	desiredTwist : Twist;
END_VAR
VAR
	speeds : WheelSpeeds;
	halfTrackInM : LREAL;
END_VAR
halfTrackInM := Parameters.trackWidthInM / 2.0;

speeds.leftInMPerS := desiredTwist.forwardSpeedInMPerS - desiredTwist.yawRateInRadPerS * halfTrackInM;
speeds.rightInMPerS := desiredTwist.forwardSpeedInMPerS + desiredTwist.yawRateInRadPerS * halfTrackInM;

ToWheelSpeeds := speeds;
END_METHOD

END_FUNCTION_BLOCK

// ---- Localization/WheelOdometry.TcPOU
{attribute 'linkalways'}
{attribute 'no_explicit_call' := 'Use the methods of this class'}
{attribute 'enable_dynamic_creation'}
FUNCTION_BLOCK WheelOdometry IMPLEMENTS I_PoseSource
VAR
	drive : I_DifferentialDrive;
	kinematics : DiffDriveKinematics;
	_pose : Pose2D;
	lastLeftInM : LREAL;
	lastRightInM : LREAL;
END_VAR

METHOD Connect
VAR_INPUT
	differentialDrive : I_DifferentialDrive;
END_VAR
drive := differentialDrive;
END_METHOD

METHOD Execute
VAR
	leftInM : LREAL;
	rightInM : LREAL;
	motion : BodyMotion;
	midHeadingInRad : LREAL;
END_VAR
leftInM := drive.LeftWheelPositionInM;
rightInM := drive.RightWheelPositionInM;

motion := kinematics.ToBodyMotion(leftDeltaInM := leftInM - lastLeftInM, rightDeltaInM := rightInM - lastRightInM);
lastLeftInM := leftInM;
lastRightInM := rightInM;

midHeadingInRad := _pose.thetaInRad + motion.headingChangeInRad / 2.0;
_pose.x := _pose.x + motion.distanceInM * COS(midHeadingInRad);
_pose.y := _pose.y + motion.distanceInM * SIN(midHeadingInRad);
_pose.thetaInRad := _pose.thetaInRad + motion.headingChangeInRad;

IF _pose.thetaInRad > PI THEN
	_pose.thetaInRad := _pose.thetaInRad - 2.0 * PI;
ELSIF _pose.thetaInRad <= -PI THEN
	_pose.thetaInRad := _pose.thetaInRad + 2.0 * PI;
END_IF
END_METHOD

PROPERTY Pose : Pose2D
GET
Pose := _pose;
END_GET
END_PROPERTY

METHOD Reset
VAR_INPUT
	pose : Pose2D;
END_VAR
_pose := pose;

lastLeftInM := drive.LeftWheelPositionInM;
lastRightInM := drive.RightWheelPositionInM;
END_METHOD

END_FUNCTION_BLOCK

// ---- Localization/GyroOdometry.TcPOU
{attribute 'linkalways'}
{attribute 'no_explicit_call' := 'Use the methods of this class'}
{attribute 'enable_dynamic_creation'}
FUNCTION_BLOCK GyroOdometry IMPLEMENTS I_PoseSource
VAR
	drive : I_DifferentialDrive;
	gyro : I_Gyro;
	kinematics : DiffDriveKinematics;
	_pose : Pose2D;
	lastLeftInM : LREAL;
	lastRightInM : LREAL;
	lastGyroTimestampInNs : ULINT;
	gyroBiasInRadPerS : LREAL;
	standStillTimer : TON;
END_VAR

METHOD Connect
VAR_INPUT
	differentialDrive : I_DifferentialDrive;
	yawGyro : I_Gyro;
END_VAR
drive := differentialDrive;
gyro := yawGyro;
END_METHOD

METHOD Execute
VAR
	leftInM : LREAL;
	rightInM : LREAL;
	motion : BodyMotion;
	midHeadingInRad : LREAL;
	headingChangeInRad : LREAL;
	dtInS : LREAL;
END_VAR
// Strekning fra hjulene
leftInM := drive.LeftWheelPositionInM;
rightInM := drive.RightWheelPositionInM;
motion := kinematics.ToBodyMotion(leftDeltaInM := leftInM - lastLeftInM, rightDeltaInM := rightInM - lastRightInM);
lastLeftInM := leftInM;
lastRightInM := rightInM;


// (rate − bias) * Parameters.gyroScale

standStillTimer(IN := drive.IsStandingStill, PT := T#500MS);
// Kursendring fra gyroen, bare når det har kommet en ny måling
IF gyro.IsValid AND gyro.TimestampInNs <> lastGyroTimestampInNs THEN
	IF gyro.TimestampInNs > lastGyroTimestampInNs THEN
		dtInS := ULINT_TO_LREAL(gyro.TimestampInNs - lastGyroTimestampInNs) * 1E-9;
	END_IF
	IF dtInS > 0 AND dtInS < 0.5 THEN
		headingChangeInRad := (gyro.YawRateInRadPerS - gyroBiasInRadPerS) * Parameters.gyroScale * dtInS;
	END_IF
	
	IF standStillTimer.Q THEN
		gyroBiasInRadPerS := gyroBiasInRadPerS + 0.01 * (gyro.YawRateInRadPerS - gyroBiasInRadPerS);
		headingChangeInRad := 0;
	END_IF
	
	lastGyroTimestampInNs := gyro.TimestampInNs;
END_IF

// Flytt roboten, med kursen midt i steget
midHeadingInRad := _pose.thetaInRad + headingChangeInRad / 2.0;
_pose.x := _pose.x + motion.distanceInM * COS(midHeadingInRad);
_pose.y := _pose.y + motion.distanceInM * SIN(midHeadingInRad);
_pose.thetaInRad := _pose.thetaInRad + headingChangeInRad;

IF _pose.thetaInRad > PI THEN
	_pose.thetaInRad := _pose.thetaInRad - 2.0 * PI;
ELSIF _pose.thetaInRad <= -PI THEN
	_pose.thetaInRad := _pose.thetaInRad + 2.0 * PI;
END_IF
END_METHOD

PROPERTY Pose : Pose2D
GET
Pose := _pose;
END_GET
END_PROPERTY

METHOD Reset
VAR_INPUT
	pose : Pose2D;
END_VAR
_pose := pose;
lastLeftInM := drive.LeftWheelPositionInM;
lastRightInM := drive.RightWheelPositionInM;
lastGyroTimestampInNs := gyro.TimestampInNs;
END_METHOD

END_FUNCTION_BLOCK

// ---- Mapping/OccupancyGrid.TcPOU
// Kartet over garasjen: et rutenett der hver rute har log-odds for at noe står der.
// 0 er ukjent, positivt er opptatt og negativt er fritt, i enheter på Constants.MAP_LOG_ODDS_PER_UNIT.
// Celle [x, y] dekker verden fra origo + (x, y) * cellestørrelse og én rute bort.
{attribute 'linkalways'}
{attribute 'no_explicit_call' := 'Use the methods of this class'}
{attribute 'enable_dynamic_creation'}
FUNCTION_BLOCK OccupancyGrid
VAR
	cells : ARRAY[0..Constants.MAP_WIDTH_IN_CELLS - 1, 0..Constants.MAP_HEIGHT_IN_CELLS - 1] OF SINT;
	_revision : UDINT;
END_VAR

// Gjør hele kartet ukjent igjen.
METHOD Clear
MEMSET(destAddr := ADR(cells), fillByte := 0, n := SIZEOF(cells));
END_METHOD

// Legger ett helt lidar-scan inn i kartet.
METHOD Integrate
VAR_IN_OUT CONSTANT
	scan : LaserScan;
END_VAR
VAR_INPUT
	// Der roboten tror den var da scannet ble ferdig.
	pose : Pose2D;
END_VAR
VAR
END_VAR
// Din oppgave (M3c). For hver stråle i fra 0 til scan.count - 1:
//  1. Hopp over stråler uten måling: rangesInM[i] er 0 når lidaren ikke fikk noe svar.
//  2. Lidaren sitter ikke nødvendigvis midt på roboten. Finn posisjonen dens i verden ved å
//     rotere (Parameters.lidarMountXInM, Parameters.lidarMountYInM) med pose.thetaInRad og
//     legge til (pose.x, pose.y).
//  3. Strålens vinkel i verden:
//     pose.thetaInRad + Parameters.lidarMountThetaInRad + scan.angleMinInRad + i * scan.angleIncrementInRad
//  4. Endepunktet er lidarposisjonen pluss avstanden langs den vinkelen (COS og SIN).
//  5. Gjør lidarposisjonen og endepunktet om til ruter med TryWorldToCell,
//     og kall TraceRay(fromCell, toCell, isHit := TRUE).
// Tenk på:
//  - Lidarens rute er den samme for alle strålene i et scan.
//  - Hva gjør du når endepunktet havner utenfor kartet?
//  - Med RPLIDAR S2E er det 1000 stråler på 10 ms. Se på Exceed-telleren i tasken når det kjører.
;
END_METHOD

// Finner ruta et punkt i verden ligger i. FALSE når punktet er utenfor kartet.
METHOD TryWorldToCell : BOOL
VAR_INPUT
	xInM : LREAL;
	yInM : LREAL;
	cell : REFERENCE TO GridCell;
END_VAR
VAR
END_VAR
// Din oppgave (M3a):
//  rute x = rundet ned ((xInM - Parameters.mapOriginXInM) / Parameters.mapCellSizeInM), og tilsvarende for y.
//  Fyll inn cell og returner TRUE bare når ruta er inne i kartet (IsInside hjelper deg).
// Pass på: LREAL_TO_DINT runder til nærmeste, og TRUNC kutter mot null. Hvilken rute havner -0.3 i da?
;
END_METHOD

// Går gjennom alle rutene fra fromCell til toCell og oppdaterer dem.
METHOD TraceRay
VAR_INPUT
	fromCell : GridCell;
	toCell : GridCell;
	// TRUE når strålen traff noe i toCell. FALSE gjør hele strålen fri, også siste rute.
	isHit : BOOL;
END_VAR
VAR
END_VAR
// Din oppgave (M3b): Bresenhams linjealgoritme.
//  - Alle rutene fra og med fromCell til (men ikke med) toCell er frie:
//    AddLogOdds(cell, Parameters.mapFreeLogOdds).
//  - toCell får AddLogOdds(toCell, Parameters.mapHitLogOdds) når isHit, ellers som en fri rute.
// Bresenham går ett steg om gangen i den retningen linja går mest, og holder rede på en
// feil-sum for å vite når den også skal ta et steg på tvers. Bare heltall, ingen COS eller SIN.
// Den må virke i alle åtte retninger: test med en stråle rett opp, rett ned, og bratt bakover.
;
END_METHOD

// Legger til log-odds i én rute og holder den innenfor ±Parameters.mapMaxLogOdds.
// Ruter utenfor kartet blir ikke rørt.
METHOD PRIVATE AddLogOdds
VAR_INPUT
	cell : GridCell;
	deltaInUnits : SINT;
END_VAR
VAR
	sum : INT;
	limit : INT;
END_VAR
IF NOT IsInside(cell) THEN
	RETURN;
END_IF
// Regn i INT, så summen ikke går rundt når SINT er full (127 + 1 blir -128).
limit := SINT_TO_INT(Parameters.mapMaxLogOdds);
sum := SINT_TO_INT(cells[cell.x, cell.y]) + SINT_TO_INT(deltaInUnits);
cells[cell.x, cell.y] := INT_TO_SINT(LIMIT(-limit, sum, limit));
END_METHOD

METHOD IsInside : BOOL
VAR_INPUT
	cell : GridCell;
END_VAR
IsInside := cell.x >= 0 AND cell.x < UINT_TO_DINT(Constants.MAP_WIDTH_IN_CELLS)
	AND cell.y >= 0 AND cell.y < UINT_TO_DINT(Constants.MAP_HEIGHT_IN_CELLS);
END_METHOD

// Log-odds i en rute, i enheter på Constants.MAP_LOG_ODDS_PER_UNIT. Ruter utenfor kartet er ukjente (0).
METHOD LogOddsAt : SINT
VAR_INPUT
	cell : GridCell;
END_VAR
IF IsInside(cell) THEN
	LogOddsAt := cells[cell.x, cell.y];
END_IF
END_METHOD

// Kopierer kartet ut til GUI-en, med et nytt revisjonsnummer.
METHOD Publish
VAR_IN_OUT
	info : MapInfo;
	target : ARRAY[0..Constants.MAP_WIDTH_IN_CELLS - 1, 0..Constants.MAP_HEIGHT_IN_CELLS - 1] OF SINT;
END_VAR
_revision := _revision + 1;
target := cells;
info.revision := _revision;
info.cellSizeInM := Parameters.mapCellSizeInM;
info.originXInM := Parameters.mapOriginXInM;
info.originYInM := Parameters.mapOriginYInM;
info.widthInCells := Constants.MAP_WIDTH_IN_CELLS;
info.heightInCells := Constants.MAP_HEIGHT_IN_CELLS;
info.logOddsPerUnit := Constants.MAP_LOG_ODDS_PER_UNIT;
END_METHOD

END_FUNCTION_BLOCK

// ---- Mission/SweepMission.TcPOU
{attribute 'linkalways'}
{attribute 'no_explicit_call' := 'Use the methods of this class'}
{attribute 'enable_dynamic_creation'}
FUNCTION_BLOCK SweepMission
VAR
	_state : MissionState := MissionState.IDLE;
	stateBeforePause : MissionState;
	lastSequence : UDINT;
	_desiredTwist : Twist;
	_hasMap : BOOL;
	requestedPose : Pose2D;
	hasPoseRequest : BOOL;
	hasMapClearRequest : BOOL;
END_VAR

METHOD Execute
IF RobotHmi.command.sequence <> lastSequence THEN
	lastSequence := RobotHmi.command.sequence;
	Handle(RobotHmi.command.code);
	RobotHmi.status.acknowledgedSequence := lastSequence;
END_IF

CASE _state OF
	MissionState.MANUAL:
		_desiredTwist := RobotHmi.command.manualTwist;
	MissionState.MAPPING:
		// Til roboten kan utforske selv (M5), kjører du den med tastaturet mens den kartlegger.
		_desiredTwist := RobotHmi.command.manualTwist;
	MissionState.SWEEPING, MissionState.RETURNING_TO_DOCK:
		// Kommer i M6: feiing og retur til lader.
		_desiredTwist := Stopped();
ELSE
	_desiredTwist := Stopped();
END_CASE

RobotHmi.status.missionState := _state;
RobotHmi.status.hasMap := _hasMap;
END_METHOD

METHOD PRIVATE Handle
VAR_INPUT
	code : HmiCommandCode;
END_VAR
RobotHmi.status.lastRejection := '';

IF code = HmiCommandCode.EMERGENCY_STOP THEN
	_state := MissionState.EMERGENCY_STOPPED;
	RETURN;
END_IF
IF code = HmiCommandCode.SET_POSE THEN
	IF IsBusy() THEN
		Reject('Stopp oppdraget før du setter posisjonen.');
	ELSE
		requestedPose := RobotHmi.command.pose;
		hasPoseRequest := TRUE;
	END_IF
	RETURN;
END_IF
IF _state = MissionState.EMERGENCY_STOPPED AND code <> HmiCommandCode.RESET THEN
	Reject('Nødstopp er aktiv. Tilbakestill først.');
	RETURN;
END_IF

CASE code OF
	HmiCommandCode.RESET:
		_state := MissionState.IDLE;
	HmiCommandCode.MANUAL_DRIVE:
		IF IsBusy() THEN
			Reject('Stopp oppdraget før du kjører manuelt.');
		ELSE
			_state := MissionState.MANUAL;
		END_IF
	HmiCommandCode.START_MAPPING:
		// Et nytt kart hver gang. Fortsetter du etter en pause, bruker du RESUME.
		_state := MissionState.MAPPING;
		_hasMap := FALSE;
		hasMapClearRequest := TRUE;
	HmiCommandCode.START_SWEEPING:
		IF _hasMap THEN
			_state := MissionState.SWEEPING;
		ELSE
			Reject('Kartet mangler. Kjør kartlegging først.');
		END_IF
	HmiCommandCode.PAUSE:
		IF IsBusy() THEN
			stateBeforePause := _state;
			_state := MissionState.PAUSED;
		ELSE
			Reject('Det er ikke noe oppdrag å pause.');
		END_IF
	HmiCommandCode.RESUME:
		IF _state = MissionState.PAUSED THEN
			_state := stateBeforePause;
		ELSE
			Reject('Det er ikke noe pauset oppdrag.');
		END_IF
	HmiCommandCode.STOP:
		IF _state = MissionState.MAPPING OR (_state = MissionState.PAUSED AND stateBeforePause = MissionState.MAPPING) THEN
			_hasMap := TRUE;
		END_IF
		_state := MissionState.IDLE;
	HmiCommandCode.GO_TO_DOCK:
		_state := MissionState.RETURNING_TO_DOCK;
END_CASE
END_METHOD

METHOD PRIVATE IsBusy : BOOL
IsBusy := _state = MissionState.MAPPING OR _state = MissionState.SWEEPING OR _state = MissionState.RETURNING_TO_DOCK;
END_METHOD

METHOD PRIVATE Reject
VAR_INPUT
	reason : STRING(80);
END_VAR
RobotHmi.status.lastRejection := reason;
END_METHOD

METHOD PRIVATE Stopped : Twist
VAR
	standingStill : Twist;
END_VAR
Stopped := standingStill;
END_METHOD

METHOD TryTakePoseRequest : BOOL
VAR_INPUT
	pose : REFERENCE TO Pose2D;
END_VAR
IF NOT hasPoseRequest THEN
	RETURN;
END_IF
pose := requestedPose;
hasPoseRequest := FALSE;
TryTakePoseRequest := TRUE;
END_METHOD

// TRUE én gang når en ny kartlegging starter, så kartet kan tømmes.
METHOD TryTakeMapClearRequest : BOOL
TryTakeMapClearRequest := hasMapClearRequest;
hasMapClearRequest := FALSE;
END_METHOD

PROPERTY State : MissionState
GET
State := _state;
END_GET
END_PROPERTY

PROPERTY DesiredTwist : Twist
GET
DesiredTwist := _desiredTwist;
END_GET
END_PROPERTY

PROPERTY ShouldDrive : BOOL
GET
ShouldDrive := _state = MissionState.MANUAL OR IsBusy();
END_GET
END_PROPERTY

END_FUNCTION_BLOCK
